FUNCTION_BLOCK FB_FolderMembers
VAR_INPUT
END_VAR
VAR_OUTPUT
END_VAR
VAR
END_VAR

PROPERTY PUBLIC Enabled : BOOL
GET // PUBLIC
END_GET
SET // PUBLIC
END_SET
END_PROPERTY

METHOD Reset : BOOL
END_METHOD

END_FUNCTION_BLOCK

(* stored: Version 1.1.0.1
   POU FB_FolderMembers: Id {04d45a1f-b0f0-4187-8258-5f6be033085c}, SpecialFunc None
   Folder Members: Id {7a43fc69-0569-41f5-b411-581f69e5d375}
   Property Enabled: Id {7b8e93e3-8545-4177-ac94-4092230dbcc1}
   Get Get: Id {4f9fa19b-92c3-4bff-a0f3-83d07b220bf7}
   Set Set: Id {4cf05f55-cfa6-43a1-b1d8-e455b26dd596}
   Method Reset: Id {b53af92c-60bb-48c4-aaa2-8bfb7cf4bdfc} *)
